// TIA Portal V20 export
Screen "SYSTEM_DIAGNOSTIC_DEVICE-VIEW"  1276x673
  ScreenItem "Title_ScreenOverview_X390_Y2" at 390,2 size 510x57  Type=HmiTextBox
  ScreenItem "Line_Header_X0_Y64" at 0,64 size 1276x0  Type=HmiLine
  ScreenItem "SysDiag_Legend" at 1185,2 size 90x60  Type=HmiButton
  ScreenItem "permanentareaborderrectangle" at 0,0 size 0x0  Type=HmiRectangle
  ScreenItem "系统诊断控制_1" at 0,66 size 1280x603  Type=HmiSystemDiagnosisControl
